Universal Robots URScript: T002_qwen2.5-coder_32b_baseline_rep2_retry2.urscript

def linear_weld_path():
    # Go to home position
    movej(get_inverse_kin([0.0, -1.823874, 1.570796, -1.570796, -1.570796, 0.0]), a=1.2, v=1.0)

    # Approach above weld start
    movel(pose_trans(get_actual_tcp_pose(), [0, 0, 50]), a=1.2, v=0.25)

    # Descend to weld start position
    movel(pose_trans(get_actual_tcp_pose(), [0, 0, -40]), a=1.2, v=0.1)

    # Weld seam — 300mm linear path
    movel(pose_trans(get_actual_tcp_pose(), [300, 0, 0]), a=1.2, v=0.05)

    # Retract above weld end
    movel(pose_trans(get_actual_tcp_pose(), [0, 0, 40]), a=1.2, v=0.2)

    # Move away from the workpiece
    movel(pose_trans(get_actual_tcp_pose(), [0, 50, 0]), a=1.2, v=0.25)
end

# Execute the weld path function
linear_weld_path()
